INTERFACE PUBLIC AsyncCommand EXTENDS Nepionic_Core.AsyncCommand

END_INTERFACE

(* stored: Version 1.1.0.1
   Itf AsyncCommand: Id {9b0fd439-a544-4026-9fa9-92113e53524a} *)
